// TIA Portal V15.1 export
ORGANIZATION_BLOCK "Main"   // OB1, LAD, ProgramCycle
TITLE = Main
{ S7_Optimized_Access := 'TRUE' }
VERSION : 0.1
// Calls the blocks in a fixed order; no logic here (decisions/0006)
// stored: AutoNumber false, IsIECCheckEnabled false, SetENOAutomatically False
   VAR_INPUT
      Initial_Call : Bool;
      Remanence : Bool;
   END_VAR
BEGIN

REGION Network 1: decisions/0006 — Common: E-STOP latch, RESET edge, parameters
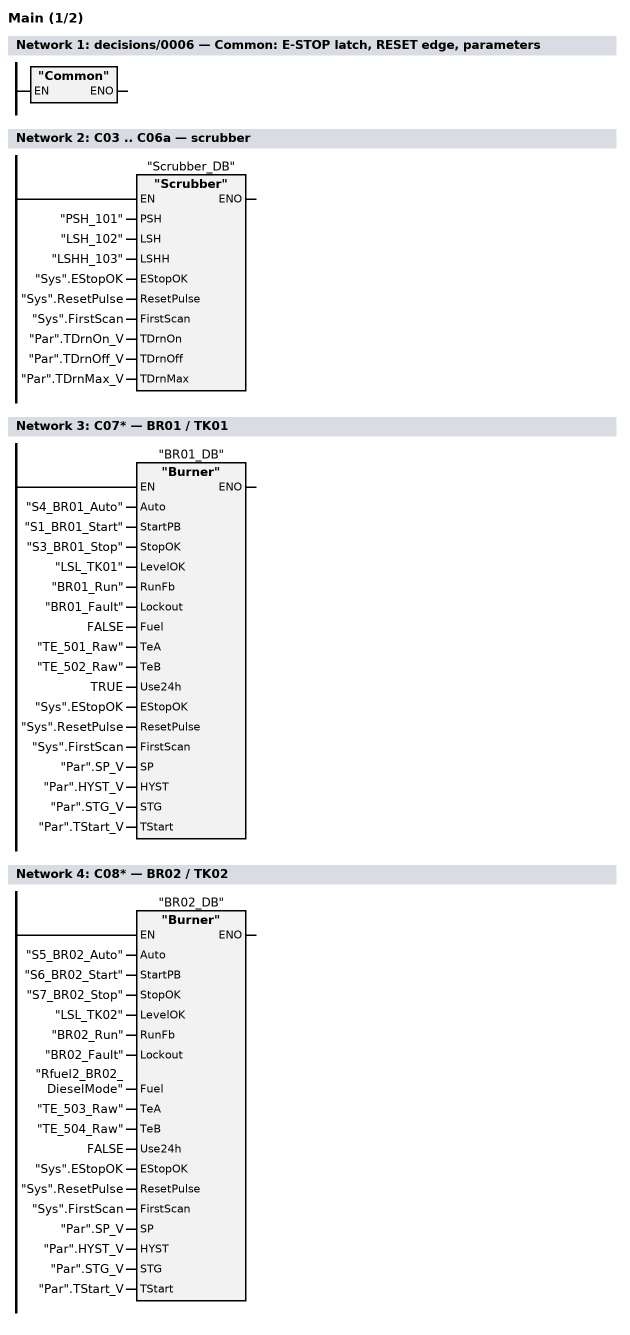
   RUNG wire#powerrail
      "Common"()
   END_RUNG
   // the same network as SCL:
   "Common"();
END_REGION

REGION Network 2: C03 .. C06a — scrubber
   RUNG wire#powerrail
      "Scrubber_DB"(PSH := "PSH_101", LSH := "LSH_102", LSHH := "LSHH_103", EStopOK := "Sys".EStopOK, ResetPulse := "Sys".ResetPulse, FirstScan := "Sys".FirstScan, TDrnOn := "Par".TDrnOn_V, TDrnOff := "Par".TDrnOff_V, TDrnMax := "Par".TDrnMax_V)
   END_RUNG
   // the same network as SCL:
   "Scrubber_DB"(PSH := "PSH_101",   // "Scrubber"
                 LSH := "LSH_102",
                 LSHH := "LSHH_103",
                 EStopOK := "Sys".EStopOK,
                 ResetPulse := "Sys".ResetPulse,
                 FirstScan := "Sys".FirstScan,
                 TDrnOn := "Par".TDrnOn_V,
                 TDrnOff := "Par".TDrnOff_V,
                 TDrnMax := "Par".TDrnMax_V);
END_REGION

REGION Network 3: C07* — BR01 / TK01
   RUNG wire#powerrail
      "BR01_DB"(Auto := "S4_BR01_Auto", StartPB := "S1_BR01_Start", StopOK := "S3_BR01_Stop", LevelOK := "LSL_TK01", RunFb := "BR01_Run", Lockout := "BR01_Fault", Fuel := FALSE, TeA := "TE_501_Raw", TeB := "TE_502_Raw", Use24h := TRUE, EStopOK := "Sys".EStopOK, ResetPulse := "Sys".ResetPulse, FirstScan := "Sys".FirstScan, SP := "Par".SP_V, HYST := "Par".HYST_V, STG := "Par".STG_V, TStart := "Par".TStart_V)
   END_RUNG
   // the same network as SCL:
   "BR01_DB"(Auto := "S4_BR01_Auto",   // "Burner"
             StartPB := "S1_BR01_Start",
             StopOK := "S3_BR01_Stop",
             LevelOK := "LSL_TK01",
             RunFb := "BR01_Run",
             Lockout := "BR01_Fault",
             Fuel := FALSE,
             TeA := "TE_501_Raw",
             TeB := "TE_502_Raw",
             Use24h := TRUE,
             EStopOK := "Sys".EStopOK,
             ResetPulse := "Sys".ResetPulse,
             FirstScan := "Sys".FirstScan,
             SP := "Par".SP_V,
             HYST := "Par".HYST_V,
             STG := "Par".STG_V,
             TStart := "Par".TStart_V);
END_REGION

REGION Network 4: C08* — BR02 / TK02
   RUNG wire#powerrail
      "BR02_DB"(Auto := "S5_BR02_Auto", StartPB := "S6_BR02_Start", StopOK := "S7_BR02_Stop", LevelOK := "LSL_TK02", RunFb := "BR02_Run", Lockout := "BR02_Fault", Fuel := "Rfuel2_BR02_DieselMode", TeA := "TE_503_Raw", TeB := "TE_504_Raw", Use24h := FALSE, EStopOK := "Sys".EStopOK, ResetPulse := "Sys".ResetPulse, FirstScan := "Sys".FirstScan, SP := "Par".SP_V, HYST := "Par".HYST_V, STG := "Par".STG_V, TStart := "Par".TStart_V)
   END_RUNG
   // the same network as SCL:
   "BR02_DB"(Auto := "S5_BR02_Auto",   // "Burner"
             StartPB := "S6_BR02_Start",
             StopOK := "S7_BR02_Stop",
             LevelOK := "LSL_TK02",
             RunFb := "BR02_Run",
             Lockout := "BR02_Fault",
             Fuel := "Rfuel2_BR02_DieselMode",
             TeA := "TE_503_Raw",
             TeB := "TE_504_Raw",
             Use24h := FALSE,
             EStopOK := "Sys".EStopOK,
             ResetPulse := "Sys".ResetPulse,
             FirstScan := "Sys".FirstScan,
             SP := "Par".SP_V,
             HYST := "Par".HYST_V,
             STG := "Par".STG_V,
             TStart := "Par".TStart_V);
END_REGION

REGION Network 5: E1 .. E7 — outputs
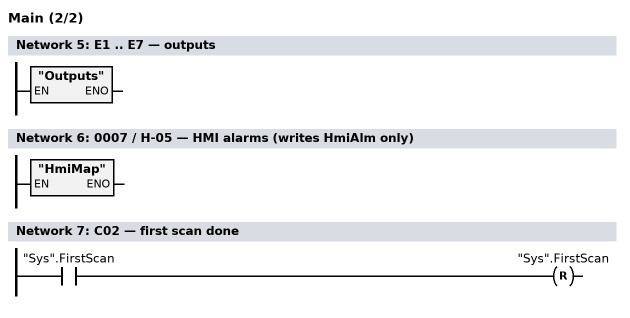
   RUNG wire#powerrail
      "Outputs"()
   END_RUNG
   // the same network as SCL:
   "Outputs"();
END_REGION

REGION Network 6: 0007 / H-05 — HMI alarms (writes HmiAlm only)
   RUNG wire#powerrail
      "HmiMap"()
   END_RUNG
   // the same network as SCL:
   "HmiMap"();
END_REGION

REGION Network 7: C02 — first scan done
   RUNG wire#powerrail
      Contact( "Sys".FirstScan )
      R_Coil( "Sys".FirstScan )
   END_RUNG
   // the same network as SCL:
   IF "Sys".FirstScan THEN "Sys".FirstScan := FALSE; END_IF;
END_REGION
END_ORGANIZATION_BLOCK
